FUNCTION_BLOCK ControlConsole (* CAT Function Block Type *)
  (* Standard: 61499-2 *)
  (* Version 0.0, 11/16/2026, Sandeep Patil, Flexbridge AB, template *)
  PACKAGE Flexbridge.FestoMPS400;
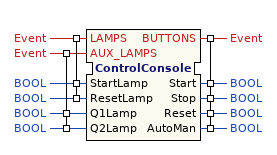
  EVENT_INPUT
    LAMPS WITH StartLamp, ResetLamp; (* START and RESET lamps (from StationMode) *)
    AUX_LAMPS WITH Q1Lamp, Q2Lamp; (* Lamps Q1 and Q2 (from the station sequence) *)
  END_EVENT
  EVENT_OUTPUT
    BUTTONS WITH Start, Stop, Reset, AutoMan; (* Button states changed *)
  END_EVENT
  VAR_INPUT
    StartLamp : BOOL; (* StartLamp on *)
    ResetLamp : BOOL; (* ResetLamp on *)
    Q1Lamp : BOOL; (* Q1Lamp on *)
    Q2Lamp : BOOL; (* Q2Lamp on *)
  END_VAR
  VAR_OUTPUT
    Start : BOOL; (* START pressed *)
    Stop : BOOL; (* STOP pressed (NC inverted) *)
    Reset : BOOL; (* RESET pressed *)
    AutoMan : BOOL; (* Key switch position *)
  END_VAR
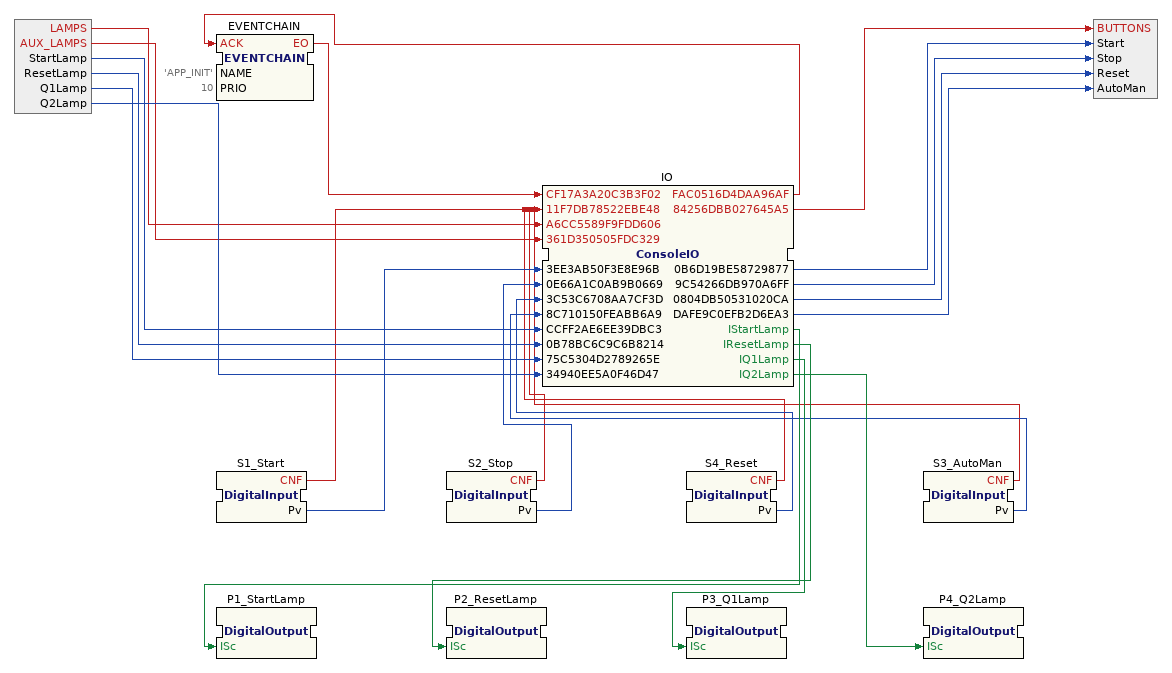
  (* 0 - INITIALIZATION *)
  (* 5 - LOGICS (ConsoleIO) *)
  (* 3.B - FROM THE FIELD (buttons, DI08-DI11) *)
  (* 3.A - TO THE FIELD (lamps, DO08-DO11) *)
  FBS
    EVENTCHAIN : EVENTCHAIN(NAME := 'APP_INIT', PRIO := 10);
    IO : ConsoleIO;
    S1_Start : DigitalInput;
    S2_Stop : DigitalInput;
    S4_Reset : DigitalInput;
    S3_AutoMan : DigitalInput;
    P1_StartLamp : DigitalOutput;
    P2_ResetLamp : DigitalOutput;
    P3_Q1Lamp : DigitalOutput;
    P4_Q2Lamp : DigitalOutput;
  END_FBS
  EVENT_CONNECTIONS
    EVENTCHAIN.EO TO IO.CF17A3A20C3B3F02;
    IO.FAC0516D4DAA96AF TO EVENTCHAIN.ACK;
    S1_Start.CNF TO IO.11F7DB78522EBE48;
    S2_Stop.CNF TO IO.11F7DB78522EBE48;
    S4_Reset.CNF TO IO.11F7DB78522EBE48;
    S3_AutoMan.CNF TO IO.11F7DB78522EBE48;
    LAMPS TO IO.A6CC5589F9FDD606;
    AUX_LAMPS TO IO.361D350505FDC329;
    IO.84256DBB027645A5 TO BUTTONS;
  END_CONNECTIONS
  DATA_CONNECTIONS
    S1_Start.Pv TO IO.3EE3AB50F3E8E96B;
    S2_Stop.Pv TO IO.0E66A1C0AB9B0669;
    S4_Reset.Pv TO IO.3C53C6708AA7CF3D;
    S3_AutoMan.Pv TO IO.8C710150FEABB6A9;
    StartLamp TO IO.CCFF2AE6EE39DBC3;
    ResetLamp TO IO.0B78BC6C9C6B8214;
    Q1Lamp TO IO.75C5304D2789265E;
    Q2Lamp TO IO.34940EE5A0F46D47;
    IO.0B6D19BE58729877 TO Start;
    IO.9C54266DB970A6FF TO Stop;
    IO.0804DB50531020CA TO Reset;
    IO.DAFE9C0EFB2D6EA3 TO AutoMan;
  END_CONNECTIONS
  ADAPTER_CONNECTIONS
    IO.IStartLamp TO P1_StartLamp.ISc;
    IO.IResetLamp TO P2_ResetLamp.ISc;
    IO.IQ1Lamp TO P3_Q1Lamp.ISc;
    IO.IQ2Lamp TO P4_Q2Lamp.ISc;
  END_CONNECTIONS
END_FUNCTION_BLOCK
